// TIA Portal project "Snap7_Variaveis" (V21)

(* hardware
DEVICE "S7-1500/ET200MP station_1"  S7-1500 station
   slot 0: "Rail_0"  Rack  6ES7 590-1***0-0AA0
   slot 0: "PM 190W 120/230VAC"  PM 190W 120/230VAC  6EP1333-4BA00
   slot 1: "PLC_1"  CPU 1516-3 PN/DP  6ES7 516-3AN01-0AB0  V2.9
      slot 3: "CPU display_1"  6ES7591-1BA00-0AA0
      slot 32768: "PROFINET interface_1"  X1
         slot 32769: "Port_1"  X1 P1
         slot 32770: "Port_2"  X1 P2
      slot 33024: "PROFINET interface_2"  X2
         slot 33025: "Port_1"  X2 P1
      slot 33280: "DP interface_1"  X3
      slot 34817: "Virtual CP interface port_1"  Virtual CP interface port  Virtual CP interface port
   slot 2: "DI 32x24VDC HF_1"  DI 32x24VDC HF  6ES7 521-1BL00-0AB0  V2.1
   slot 3: "DQ 32x24VDC/0.5A HF_1"  DQ 32x24VDC/0.5A HF  6ES7 522-1BL01-0AB0  V1.0
   slot 4: "AI 8xU/I/RTD/TC ST_1"  AI 8xU/I/RTD/TC ST  6ES7 531-7KF00-0AB0  V2.0
   slot 5: "AQ 4xU/I ST_1"  AQ 4xU/I ST  6ES7 532-5HD00-0AB0  V2.0
*)

// ===== PLC "PLC_1"  CPU 1516-3 PN/DP =====

DATA_BLOCK "DB_Snap7"   // DB1
{ S7_Optimized_Access := 'FALSE' }
   VAR
      Bool_0 : Bool;
      Bool_1 : Bool;
      Bool_2 : Bool;
      Bool_3 : Bool;
      Bool_4 : Bool;
      Bool_5 : Bool;
      Bool_6 : Bool;
      Bool_7 : Bool;
      Byte_Val : Byte;
      Int_Val : Int;
      UInt_Val : UInt;
      Word_Val : Word;
      LReal_Val : LReal;
      DInt_Val : DInt;
      UDInt_Val : UDInt;
      Real_Val : Real;
      String_Val : String[20];
      SInt_Val : SInt;
      USInt_Val : USInt;
   END_VAR
BEGIN
END_DATA_BLOCK

DATA_BLOCK "DB_Snap7_Resp"   // DB2
{ S7_Optimized_Access := 'FALSE' }
   VAR
      Heartbeat : Bool;
      E_Bool01 : Bool;
      OU_Bool23 : Bool;
      NAO_Bool4 : Bool;
      Qualquer_Bool : Bool;
      Soma_Bits : Byte;
      Int_Mais1 : Int;
      DInt_Dobro : DInt;
      Contador : DInt;
      Real_Fahrenheit : Real;
      LReal_Raiz : LReal;
      String_Eco : String[30];
      Len_String : Int;
      Word_Invertida : Word;
      tmrContador : TON_TIME;
      tmrHeartbeat : TON_TIME;
   END_VAR
BEGIN
END_DATA_BLOCK

DATA_BLOCK "DB_Snap7_Aux"   // DB3
{ S7_Optimized_Access := 'FALSE' }
   VAR
      UltTickContador : DInt;
      UltTickHeartbeat : DInt;
   END_VAR
BEGIN
END_DATA_BLOCK

FUNCTION "FC_Logica_Snap7" : Void   // FC1, SCL
{ S7_Optimized_Access := 'TRUE' }
VERSION : 0.2
   VAR_TEMP
      soma : USInt;
      agora : DInt;
      dif : DInt;
   END_VAR
BEGIN

       // Entradas: DB_Snap7 (escritas pelo Python via Snap7)
       // Saidas:   DB_Snap7_Resp (calculadas aqui, lidas pelo Python)
       // Bool_6 = pausa o contador | Bool_7 = zera o contador
       // Tempo: comparacao com o relogio da CPU (TIME_TCK), sem timers IEC

       // ---- Bool ----
       "DB_Snap7_Resp".E_Bool01 := "DB_Snap7".Bool_0 AND "DB_Snap7".Bool_1;
       "DB_Snap7_Resp".OU_Bool23 := "DB_Snap7".Bool_2 OR "DB_Snap7".Bool_3;
       "DB_Snap7_Resp".NAO_Bool4 := NOT "DB_Snap7".Bool_4;

       #soma := 0;
       IF "DB_Snap7".Bool_0 THEN #soma := #soma + 1; END_IF;
       IF "DB_Snap7".Bool_1 THEN #soma := #soma + 1; END_IF;
       IF "DB_Snap7".Bool_2 THEN #soma := #soma + 1; END_IF;
       IF "DB_Snap7".Bool_3 THEN #soma := #soma + 1; END_IF;
       IF "DB_Snap7".Bool_4 THEN #soma := #soma + 1; END_IF;
       IF "DB_Snap7".Bool_5 THEN #soma := #soma + 1; END_IF;
       IF "DB_Snap7".Bool_6 THEN #soma := #soma + 1; END_IF;
       IF "DB_Snap7".Bool_7 THEN #soma := #soma + 1; END_IF;
       "DB_Snap7_Resp".Soma_Bits := USINT_TO_BYTE(#soma);
       "DB_Snap7_Resp".Qualquer_Bool := #soma > 0;

       // ---- Inteiros ----
       IF "DB_Snap7".Int_Val < 32767 THEN
           "DB_Snap7_Resp".Int_Mais1 := "DB_Snap7".Int_Val + 1;
       ELSE
           "DB_Snap7_Resp".Int_Mais1 := 32767;
       END_IF;
       "DB_Snap7_Resp".DInt_Dobro := INT_TO_DINT("DB_Snap7".Int_Val) * 2;

       // ---- Reais ----
       "DB_Snap7_Resp".Real_Fahrenheit := "DB_Snap7".Real_Val * 1.8 + 32.0;
       "DB_Snap7_Resp".LReal_Raiz := SQRT(ABS("DB_Snap7".LReal_Val));

       // ---- String / Word ----
       "DB_Snap7_Resp".String_Eco := CONCAT(IN1 := 'Eco: ', IN2 := "DB_Snap7".String_Val);
       "DB_Snap7_Resp".Len_String := LEN("DB_Snap7".String_Val);
       "DB_Snap7_Resp".Word_Invertida := NOT "DB_Snap7".Word_Val;

       // ---- Tempo atual da CPU em ms ----
       #agora := TIME_TO_DINT(TIME_TCK());

       // ---- Contador (+1 a cada 100 ms) ----
       #dif := #agora - "DB_Snap7_Aux".UltTickContador;
       IF (#dif >= 100) OR (#dif < 0) THEN
           "DB_Snap7_Aux".UltTickContador := #agora;
           IF NOT "DB_Snap7".Bool_6 THEN
               IF "DB_Snap7_Resp".Contador < 2147483647 THEN
                   "DB_Snap7_Resp".Contador := "DB_Snap7_Resp".Contador + 1;
               END_IF;
           END_IF;
       END_IF;
       IF "DB_Snap7".Bool_7 THEN
           "DB_Snap7_Resp".Contador := 0;
       END_IF;

       // ---- Heartbeat (alterna a cada 500 ms) ----
       #dif := #agora - "DB_Snap7_Aux".UltTickHeartbeat;
       IF (#dif >= 500) OR (#dif < 0) THEN
           "DB_Snap7_Aux".UltTickHeartbeat := #agora;
           "DB_Snap7_Resp".Heartbeat := NOT "DB_Snap7_Resp".Heartbeat;
       END_IF;
END_FUNCTION

ORGANIZATION_BLOCK "Main"   // OB1, LAD, ProgramCycle
TITLE = "Main Program Sweep (Cycle)"
{ S7_Optimized_Access := 'TRUE' }
VERSION : 0.1
   VAR_INPUT
      Initial_Call : Bool;   // Initial call of this OB
      Remanence : Bool;   // =True, if remanent data are available
   END_VAR
BEGIN

REGION Network 1
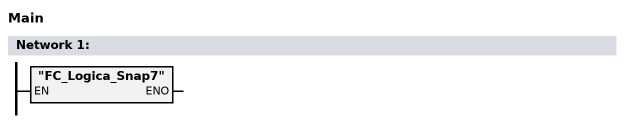
   RUNG wire#powerrail
      "FC_Logica_Snap7"()
   END_RUNG
   // the same network as SCL:
   "FC_Logica_Snap7"();
END_REGION
END_ORGANIZATION_BLOCK